{attribute 'linkalways'} 
{attribute 'no_explicit_call' := 'This FB is a CLASS and must be accessed using methods or properties'}
{attribute 'enable_dynamic_creation'}
FUNCTION_BLOCK _Array0to3OfSINT EXTENDS ArrayDatatypeBase_1D
VAR CONSTANT
	lBound : DINT := 0;
	uBound : DINT := 3;
END_VAR
VAR
	localData : ARRAY [lBound..uBound] OF SINT;
	activeData : REFERENCE TO ARRAY [lBound..uBound] OF SINT REF= localData;
	elements : ARRAY [lBound..uBound] OF _SINT(0);
	baseType : _SINT(0);
END_VAR

PROPERTY PUBLIC Address : PVOID
GET
Address := ADR(activeData);
END_GET
END_PROPERTY

PROPERTY PUBLIC BaseDatatype : I_Datatype
GET
BaseDatatype := baseType;
END_GET
END_PROPERTY

METHOD PUBLIC ClearReference
VAR_INPUT
END_VAR
activeData REF= localData;
SetElementReference();
END_METHOD

METHOD PUBLIC Clone : I_Datatype
VAR
    pClone : POINTER TO _Array0to3OfSINT;
END_VAR
pClone := __NEW(_Array0to3OfSINT());
pClone^.Value := Value;
Clone := pClone^;
END_METHOD

METHOD FB_init : BOOL
VAR_INPUT
	bInitRetains : BOOL; // if TRUE, the retain variables are initialized (warm start / cold start)
	bInCopyCode : BOOL;  // if TRUE, the instance afterwards gets moved into the copy code (online change)
END_VAR
SetElementReference();
END_METHOD

METHOD PUBLIC MakeReferenceTo
VAR_INPUT
	ReferenceTarget : REFERENCE TO ARRAY [lBound..uBound] OF SINT;
END_VAR
activeData REF= ReferenceTarget;
SetElementReference();
END_METHOD

METHOD PROTECTED OnSerializeArrayValues
VAR_INPUT
	Serializer : I_Serializer;
END_VAR
VAR
	i : DINT;
END_VAR
FOR i := lBound TO uBound DO
	elements[i].SerializeWith(Serializer);
END_FOR
END_METHOD

METHOD PROTECTED SetElementReference
VAR_INPUT
END_VAR
VAR
	i : DINT;
END_VAR
FOR i := lBound TO uBound DO
	elements[i].MakeReferenceTo(activeData[i]);
END_FOR
END_METHOD

PROPERTY PUBLIC Size : UDINT
GET
Size := SIZEOF(activeData);
END_GET
END_PROPERTY

METHOD PROTECTED TryDeserializeArrayValues : BOOL
VAR_INPUT
	Deserializer : I_Deserializer;
	Feedback : I_DeserializerFeedback;
END_VAR
VAR
	failed : BOOL;
	enumerator : I_DeserializerArrayForwardEnumerator;
	i : DINT;
END_VAR
enumerator := Deserializer.GetArrayEnumerator();
i := lBound;

WHILE enumerator.MoveNext() AND i <= uBound AND NOT failed DO
	
	IF NOT elements[i].TryDeserializeFrom(enumerator.Current, Feedback) THEN
		failed := TRUE;
		EXIT;
	END_IF
	i := i + 1;

END_WHILE
enumerator.Dispose();

TryDeserializeArrayValues := NOT failed;
END_METHOD

METHOD PUBLIC TryGetElementAsDatatypeByIndex : BOOL
VAR_INPUT
	Index : DINT;
	Destination : REFERENCE TO I_Datatype;
END_VAR
IF Index < lbound OR Index > ubound THEN
	RETURN;
END_IF

Destination := elements[Index];
TryGetElementAsDatatypeByIndex := TRUE;
END_METHOD

METHOD PUBLIC TryGetLowerBound : BOOL
VAR_INPUT
	Dimention : UDINT;
	Destination : REFERENCE TO DINT;
END_VAR
IF Dimention = 1 THEN
	Destination := lBound;
	TryGetLowerBound := TRUE;
END_IF
END_METHOD

METHOD PUBLIC TryGetUpperBound : BOOL
VAR_INPUT
	Dimention : UDINT;
	Destination : REFERENCE TO DINT;
END_VAR
IF Dimention = 1 THEN
	Destination := uBound;
	TryGetUpperBound := TRUE;
END_IF
END_METHOD

METHOD TryMakeReferenceTo : BOOL
VAR_INPUT
	Target : I_Datatype;
END_VAR
VAR
	pTargetData : POINTER TO ARRAY [lBound..uBound] OF SINT;
END_VAR
IF NOT IsEquivalentTo(Target) THEN
	RETURN;
END_IF

pTargetData := Target.Address;
activeData REF= pTargetData^;
SetElementReference();
TryMakeReferenceTo := TRUE;
END_METHOD

PROPERTY PUBLIC Value : REFERENCE TO ARRAY [lBound..uBound] OF SINT;
GET
Value ref= activeData;
END_GET
END_PROPERTY

END_FUNCTION_BLOCK

(* stored: Version 1.1.0.1, ProductVersion 3.1.4024.13
   POU _Array0to3OfSINT: Id {872bbb7b-8a04-0a2b-0db3-20bc2659623d}, SpecialFunc None
   Folder Core: Id {c89e7023-eb0d-0a76-3d39-60a5711def5e}
   Folder Constructor: Id {e94fce87-bbd5-0ae4-026e-ed50b08c4f80}
   Folder Protected: Id {aaf18fb3-7346-0ae6-16df-754456ef7d5e}
   Folder Customize: Id {1449433a-50ba-0c1f-14d6-31e3878aaa81}
   Property Address: Id {8174a0c9-99ab-01b0-3b3e-a0e6a764dfc7}
   Get Get: Id {cae941d0-f6a2-02d9-10e0-2d82caf72b4a}
   Property BaseDatatype: Id {c12a4a09-b2d9-03a5-082c-1cf529158bcc}
   Get Get: Id {073f37c3-bc99-01b4-3d99-6fee074153d8}
   Method ClearReference: Id {81865733-ebbb-053d-1aef-bf17bb685624}
   Method Clone: Id {dc19fcdb-ca23-076c-14d0-c54bcc61a6f0}
   Method FB_init: Id {7c304e62-ade9-09b7-016f-ee172548defc}
   Method MakeReferenceTo: Id {4272f35b-3770-058e-3fdc-0c4f09105710}
   Method OnSerializeArrayValues: Id {3be195a7-ffc6-0d71-00a3-14ad90283271}
   Method SetElementReference: Id {5a2b0916-91c3-0def-1a76-6ea3a918c459}
   Property Size: Id {10f7e279-cc23-0d7f-0eef-7911bb6751f8}
   Get Get: Id {0cec377f-b8da-02cf-16ae-f84ad4bddad1}
   Method TryDeserializeArrayValues: Id {7ad20c17-5c36-0afd-32d2-f5d522d1d82f}
   Method TryGetElementAsDatatypeByIndex: Id {0147fff8-b90c-0ee5-3c77-054fea214c05}
   Method TryGetLowerBound: Id {6231b67b-a0da-0ed5-1335-4e77e30e2058}
   Method TryGetUpperBound: Id {79bd229c-d625-01a7-30e6-cc7833209e2c}
   Method TryMakeReferenceTo: Id {74cf5e69-17b9-0546-223d-45c29df781ed}
   Property Value: Id {652e022f-b9e1-0ff6-1e10-5f110fd1c75c}
   Get Get: Id {5a946149-54c9-01a0-3a92-58c115d6f499} *)
